// TIA Portal V20 export
// export: Created 2026-10-12T05:00:33.5810013Z, ExportSetting WithDefaults, DisplayName Totally Integrated Automation Portal, DisplayVersion V20, DisplayName TIA Portal Openness, DisplayVersion V20, DisplayName TIA Portal Teamcenter Gateway, DisplayVersion V20, DisplayName TIA Portal Version Control Interface, DisplayVersion V20, DisplayName SINAMICS Startdrive Advanced, DisplayVersion V20 SP1 Update 2, DisplayName SINAMICS Startdrive G110M, G120, G120C, G120D, G120P, G115D, DisplayVersion V20 SP1 Update 2, DisplayName SINAMICS Startdrive G130, G150, S120, S150, SINAMICS MV, G220, S200, S210, DisplayVersion V20 SP1 Update 2, DisplayName STEP 7 Professional, DisplayVersion V20, DisplayName STEP 7 Safety, DisplayVersion V20, DisplayName WinCC Basic/Comfort/Advanced, DisplayVersion V20, DisplayName WinCC Professional, DisplayVersion V20, DisplayName WinCC Unified, DisplayVersion V20
FUNCTION "F_AccessBenchProvision" : Void   // FC168, SCL
{ S7_Optimized_Access := 'TRUE' }
VERSION : 0.1
// stored: AutoNumber true, IsIECCheckEnabled false, SetENOAutomatically false, UDAEnableTagReadback false
BEGIN

   "FRK_LocalUsers".Count := 2;
   "FRK_LocalUsers".Rows[1].User := 'operator';
   "FRK_LocalUsers".Rows[1].Level := 1;
   "FRK_LocalUsers".Rows[1].Salt[0] := BYTE#16#29;
   "FRK_LocalUsers".Rows[1].Salt[1] := BYTE#16#7B;
   "FRK_LocalUsers".Rows[1].Salt[2] := BYTE#16#70;
   "FRK_LocalUsers".Rows[1].Salt[3] := BYTE#16#0D;
   "FRK_LocalUsers".Rows[1].Salt[4] := BYTE#16#96;
   "FRK_LocalUsers".Rows[1].Salt[5] := BYTE#16#3A;
   "FRK_LocalUsers".Rows[1].Salt[6] := BYTE#16#CC;
   "FRK_LocalUsers".Rows[1].Salt[7] := BYTE#16#D0;
   "FRK_LocalUsers".Rows[1].Salt[8] := BYTE#16#8A;
   "FRK_LocalUsers".Rows[1].Salt[9] := BYTE#16#25;
   "FRK_LocalUsers".Rows[1].Salt[10] := BYTE#16#55;
   "FRK_LocalUsers".Rows[1].Salt[11] := BYTE#16#F5;
   "FRK_LocalUsers".Rows[1].Salt[12] := BYTE#16#51;
   "FRK_LocalUsers".Rows[1].Salt[13] := BYTE#16#71;
   "FRK_LocalUsers".Rows[1].Salt[14] := BYTE#16#D6;
   "FRK_LocalUsers".Rows[1].Salt[15] := BYTE#16#A8;
   "FRK_LocalUsers".Rows[1].PinHash[0] := BYTE#16#96;
   "FRK_LocalUsers".Rows[1].PinHash[1] := BYTE#16#3E;
   "FRK_LocalUsers".Rows[1].PinHash[2] := BYTE#16#4A;
   "FRK_LocalUsers".Rows[1].PinHash[3] := BYTE#16#A4;
   "FRK_LocalUsers".Rows[1].PinHash[4] := BYTE#16#E0;
   "FRK_LocalUsers".Rows[1].PinHash[5] := BYTE#16#8E;
   "FRK_LocalUsers".Rows[1].PinHash[6] := BYTE#16#33;
   "FRK_LocalUsers".Rows[1].PinHash[7] := BYTE#16#94;
   "FRK_LocalUsers".Rows[1].PinHash[8] := BYTE#16#83;
   "FRK_LocalUsers".Rows[1].PinHash[9] := BYTE#16#FD;
   "FRK_LocalUsers".Rows[1].PinHash[10] := BYTE#16#D1;
   "FRK_LocalUsers".Rows[1].PinHash[11] := BYTE#16#A7;
   "FRK_LocalUsers".Rows[1].PinHash[12] := BYTE#16#CF;
   "FRK_LocalUsers".Rows[1].PinHash[13] := BYTE#16#65;
   "FRK_LocalUsers".Rows[1].PinHash[14] := BYTE#16#A6;
   "FRK_LocalUsers".Rows[1].PinHash[15] := BYTE#16#71;
   "FRK_LocalUsers".Rows[1].PinHash[16] := BYTE#16#7E;
   "FRK_LocalUsers".Rows[1].PinHash[17] := BYTE#16#29;
   "FRK_LocalUsers".Rows[1].PinHash[18] := BYTE#16#FD;
   "FRK_LocalUsers".Rows[1].PinHash[19] := BYTE#16#87;
   "FRK_LocalUsers".Rows[1].PinHash[20] := BYTE#16#37;
   "FRK_LocalUsers".Rows[1].PinHash[21] := BYTE#16#8F;
   "FRK_LocalUsers".Rows[1].PinHash[22] := BYTE#16#20;
   "FRK_LocalUsers".Rows[1].PinHash[23] := BYTE#16#B0;
   "FRK_LocalUsers".Rows[1].PinHash[24] := BYTE#16#DC;
   "FRK_LocalUsers".Rows[1].PinHash[25] := BYTE#16#A6;
   "FRK_LocalUsers".Rows[1].PinHash[26] := BYTE#16#7B;
   "FRK_LocalUsers".Rows[1].PinHash[27] := BYTE#16#1F;
   "FRK_LocalUsers".Rows[1].PinHash[28] := BYTE#16#0B;
   "FRK_LocalUsers".Rows[1].PinHash[29] := BYTE#16#51;
   "FRK_LocalUsers".Rows[1].PinHash[30] := BYTE#16#64;
   "FRK_LocalUsers".Rows[1].PinHash[31] := BYTE#16#0B;
   "FRK_LocalUsers".Rows[2].User := 'admin';
   "FRK_LocalUsers".Rows[2].Level := 4;
   "FRK_LocalUsers".Rows[2].Salt[0] := BYTE#16#5A;
   "FRK_LocalUsers".Rows[2].Salt[1] := BYTE#16#41;
   "FRK_LocalUsers".Rows[2].Salt[2] := BYTE#16#72;
   "FRK_LocalUsers".Rows[2].Salt[3] := BYTE#16#AC;
   "FRK_LocalUsers".Rows[2].Salt[4] := BYTE#16#00;
   "FRK_LocalUsers".Rows[2].Salt[5] := BYTE#16#2B;
   "FRK_LocalUsers".Rows[2].Salt[6] := BYTE#16#38;
   "FRK_LocalUsers".Rows[2].Salt[7] := BYTE#16#55;
   "FRK_LocalUsers".Rows[2].Salt[8] := BYTE#16#53;
   "FRK_LocalUsers".Rows[2].Salt[9] := BYTE#16#4A;
   "FRK_LocalUsers".Rows[2].Salt[10] := BYTE#16#AE;
   "FRK_LocalUsers".Rows[2].Salt[11] := BYTE#16#0E;
   "FRK_LocalUsers".Rows[2].Salt[12] := BYTE#16#0C;
   "FRK_LocalUsers".Rows[2].Salt[13] := BYTE#16#C9;
   "FRK_LocalUsers".Rows[2].Salt[14] := BYTE#16#F6;
   "FRK_LocalUsers".Rows[2].Salt[15] := BYTE#16#9C;
   "FRK_LocalUsers".Rows[2].PinHash[0] := BYTE#16#FA;
   "FRK_LocalUsers".Rows[2].PinHash[1] := BYTE#16#3F;
   "FRK_LocalUsers".Rows[2].PinHash[2] := BYTE#16#3C;
   "FRK_LocalUsers".Rows[2].PinHash[3] := BYTE#16#F5;
   "FRK_LocalUsers".Rows[2].PinHash[4] := BYTE#16#C0;
   "FRK_LocalUsers".Rows[2].PinHash[5] := BYTE#16#79;
   "FRK_LocalUsers".Rows[2].PinHash[6] := BYTE#16#91;
   "FRK_LocalUsers".Rows[2].PinHash[7] := BYTE#16#CF;
   "FRK_LocalUsers".Rows[2].PinHash[8] := BYTE#16#1D;
   "FRK_LocalUsers".Rows[2].PinHash[9] := BYTE#16#81;
   "FRK_LocalUsers".Rows[2].PinHash[10] := BYTE#16#BD;
   "FRK_LocalUsers".Rows[2].PinHash[11] := BYTE#16#8C;
   "FRK_LocalUsers".Rows[2].PinHash[12] := BYTE#16#66;
   "FRK_LocalUsers".Rows[2].PinHash[13] := BYTE#16#AA;
   "FRK_LocalUsers".Rows[2].PinHash[14] := BYTE#16#90;
   "FRK_LocalUsers".Rows[2].PinHash[15] := BYTE#16#E5;
   "FRK_LocalUsers".Rows[2].PinHash[16] := BYTE#16#82;
   "FRK_LocalUsers".Rows[2].PinHash[17] := BYTE#16#E1;
   "FRK_LocalUsers".Rows[2].PinHash[18] := BYTE#16#CB;
   "FRK_LocalUsers".Rows[2].PinHash[19] := BYTE#16#81;
   "FRK_LocalUsers".Rows[2].PinHash[20] := BYTE#16#9D;
   "FRK_LocalUsers".Rows[2].PinHash[21] := BYTE#16#52;
   "FRK_LocalUsers".Rows[2].PinHash[22] := BYTE#16#77;
   "FRK_LocalUsers".Rows[2].PinHash[23] := BYTE#16#75;
   "FRK_LocalUsers".Rows[2].PinHash[24] := BYTE#16#3B;
   "FRK_LocalUsers".Rows[2].PinHash[25] := BYTE#16#30;
   "FRK_LocalUsers".Rows[2].PinHash[26] := BYTE#16#88;
   "FRK_LocalUsers".Rows[2].PinHash[27] := BYTE#16#8F;
   "FRK_LocalUsers".Rows[2].PinHash[28] := BYTE#16#7F;
   "FRK_LocalUsers".Rows[2].PinHash[29] := BYTE#16#15;
   "FRK_LocalUsers".Rows[2].PinHash[30] := BYTE#16#DA;
   "FRK_LocalUsers".Rows[2].PinHash[31] := BYTE#16#44;

   "GDB_AccessPersistTest".ProvisionCount := "GDB_AccessPersistTest".ProvisionCount + 1;
END_FUNCTION
